TYPE "ST_DataClassPolicy"
VERSION : 0.1
   STRUCT
      ClassId : String[40];
      LabelKey : String[160];
      ReadLevel : DInt;
      WriteLevel : DInt;
   END_STRUCT;

END_TYPE

